Fanuc KAREL source: NC0051.KL

-- PROVISIONAL review KL for V770-1; original PC SHA256 e07c157cf1558a2f99da5237d425802c3457d570def0ff00f2ca9d62f1d1d3d1
-- Incomplete behavior may be omitted. Consult companion uncertainty JSON. Do not deploy.
PROGRAM NC0051
%NOLOCKGROUP
-- UNRESOLVED_LOCAL_POOL 1 cells at code offset 3; source declarations unknown
-- DIRECT_LOCAL_WORD_ACCESS alone does not prove INTEGER, REAL, or BOOLEAN
BEGIN
  -- UNRESOLVED_PC offsets 0-8; opcodes 2B,2C,7B
  -- UNRESOLVED_PC offsets 13-20; opcodes 9D,23
  -- UNRESOLVED_PC offsets 25-38; opcodes 21,9D,57,79
  -- UNRESOLVED_PC offsets 43-60; opcodes 21,40,41,42
  -- UNRESOLVED_PC offsets 65-78; opcodes 21,9D,57,79
  -- UNRESOLVED_PC offsets 83-100; opcodes 21,40,41,42
  -- UNRESOLVED_PC offsets 105-118; opcodes 21,9D,57,79
  -- UNRESOLVED_PC offsets 123-140; opcodes 21,40,41,42
  -- UNRESOLVED_PC offsets 145-158; opcodes 21,9D,57,79
  -- UNRESOLVED_PC offsets 163-180; opcodes 21,40,41,42
  -- UNRESOLVED_PC offsets 185-198; opcodes 21,9D,57,79
  -- UNRESOLVED_PC offsets 203-220; opcodes 21,40,41,42
  -- UNRESOLVED_PC offsets 225-238; opcodes 21,9D,57,79
  -- UNRESOLVED_PC offsets 243-260; opcodes 21,40,41,42
  -- UNRESOLVED_PC offsets 265-278; opcodes 21,9D,57,79
  -- UNRESOLVED_PC offsets 283-300; opcodes 21,40,41,42
  -- UNRESOLVED_PC offsets 305-318; opcodes 21,9D,57,79
  -- UNRESOLVED_PC offsets 323-340; opcodes 21,40,41,42
  -- UNRESOLVED_PC offsets 345-358; opcodes 21,9D,57,79
  -- UNRESOLVED_PC offsets 363-380; opcodes 21,40,41,42
  -- UNRESOLVED_PC offsets 385-398; opcodes 21,9D,57,79
  -- UNRESOLVED_PC offsets 403-420; opcodes 21,40,41,42
  -- UNRESOLVED_PC offsets 425-455; opcodes 21,9D,52,23,7A,40,41,42
  -- UNRESOLVED_PC offsets 460-484; opcodes 21,2E,52,23,7A,43
  -- UNRESOLVED_PC offsets 489-507; opcodes 21,2E,52,23
  -- UNRESOLVED_PC offsets 517-522; opcodes 7A
  -- UNRESOLVED_PC offsets 527-545; opcodes 21,2E,52,23
  -- UNRESOLVED_PC offsets 550-566; opcodes 7A,40,41,42
  -- UNRESOLVED_PC offsets 571-595; opcodes 21,2E,52,23,7A,43
  -- UNRESOLVED_PC offsets 600-618; opcodes 21,2E,52,23
  -- UNRESOLVED_PC offsets 628-633; opcodes 7A
  -- UNRESOLVED_PC offsets 638-656; opcodes 21,2E,52,23
  -- UNRESOLVED_PC offsets 661-677; opcodes 7A,40,41,42
  -- UNRESOLVED_PC offsets 682-706; opcodes 21,2E,52,23,7A,43
  -- UNRESOLVED_PC offsets 711-729; opcodes 21,2E,52,23
  -- UNRESOLVED_PC offsets 739-744; opcodes 7A
  -- UNRESOLVED_PC offsets 749-767; opcodes 21,2E,52,23
  -- UNRESOLVED_PC offsets 772-788; opcodes 7A,40,41,42
  -- UNRESOLVED_PC offsets 793-817; opcodes 21,2E,52,23,7A,43
  -- UNRESOLVED_PC offsets 822-840; opcodes 21,2E,52,23
  -- UNRESOLVED_PC offsets 850-855; opcodes 7A
  -- UNRESOLVED_PC offsets 860-878; opcodes 21,2E,52,23
  -- UNRESOLVED_PC offsets 883-899; opcodes 7A,40,41,42
  -- UNRESOLVED_PC offsets 904-928; opcodes 21,2E,52,23,7A,43
  -- UNRESOLVED_PC offsets 933-951; opcodes 21,2E,52,23
  -- UNRESOLVED_PC offsets 961-966; opcodes 7A
  -- UNRESOLVED_PC offsets 971-989; opcodes 21,2E,52,23
  -- UNRESOLVED_PC offsets 994-1010; opcodes 7A,40,41,42
  -- UNRESOLVED_PC offsets 1015-1039; opcodes 21,2E,52,23,7A,43
  -- UNRESOLVED_PC offsets 1044-1062; opcodes 21,2E,52,23
  -- UNRESOLVED_PC offsets 1072-1077; opcodes 7A
  -- UNRESOLVED_PC offsets 1082-1100; opcodes 21,2E,52,23
  -- UNRESOLVED_PC offsets 1105-1121; opcodes 7A,40,41,42
  -- UNRESOLVED_PC offsets 1126-1150; opcodes 21,2E,52,23,7A,43
  -- UNRESOLVED_PC offsets 1155-1173; opcodes 21,2E,52,23
  -- UNRESOLVED_PC offsets 1183-1188; opcodes 7A
  -- UNRESOLVED_PC offsets 1193-1211; opcodes 21,2E,52,23
  -- UNRESOLVED_PC offsets 1216-1232; opcodes 7A,40,41,42
  -- UNRESOLVED_PC offsets 1237-1261; opcodes 21,2E,52,23,7A,43
  -- UNRESOLVED_PC offsets 1266-1284; opcodes 21,2E,52,23
  -- UNRESOLVED_PC offsets 1294-1299; opcodes 7A
  -- UNRESOLVED_PC offsets 1304-1322; opcodes 21,2E,52,23
  -- UNRESOLVED_PC offsets 1327-1343; opcodes 7A,40,41,42
  -- UNRESOLVED_PC offsets 1348-1372; opcodes 21,2E,52,23,7A,43
  -- UNRESOLVED_PC offsets 1377-1395; opcodes 21,2E,52,23
  -- UNRESOLVED_PC offsets 1405-1410; opcodes 7A
  -- UNRESOLVED_PC offsets 1415-1433; opcodes 21,2E,52,23
  -- UNRESOLVED_PC offsets 1438-1454; opcodes 7A,40,41,42
  -- UNRESOLVED_PC offsets 1459-1483; opcodes 21,2E,52,23,7A,43
  -- UNRESOLVED_PC offsets 1488-1506; opcodes 21,2E,52,23
  -- UNRESOLVED_PC offsets 1516-1521; opcodes 7A
  -- UNRESOLVED_PC offsets 1526-1544; opcodes 21,2E,52,23
  -- UNRESOLVED_PC offsets 1554-1558; opcodes 7F
  -- UNRESOLVED_PC offsets 1563-1567; opcodes 27,AA
  -- UNRESOLVED_PC offsets 1572-1576; opcodes 7F
END NC0051
